(* IEC 61131-3 sources: iolistgen/tools/tests/fixtures/sample/tests/POUs/PRG_Tests, 1 file *)

(* ---- PRG_Tests.decl.st ---- *)
(*
    Назначение: запуск тестов CfUnit
    Автор: kr0nsch
    Версия: 1.0.0
    Документ: docs/TEST_REPORT.md
*)
PROGRAM PRG_Tests
VAR
    fbClampTest : FB_F_Clamp_Test;
END_VAR
